(* IEC 61131-3 sources: nautilus/examples/remote-fleet/scada, 2 files *)

(* ---- sparkplug_types.st ---- *)
(*
  Generated by `naut sparkplug import` from the group's NBIRTH template
  definitions. Do not edit — re-run the import when a site's UDTs change.
  Group: Water
*)

TYPE
  Pump : STRUCT
    Run : BOOL;
    Fault : BOOL;
    SpeedHz : LREAL;
    SpeedSP : LREAL;
  END_STRUCT;
END_TYPE

(* Add the tags your program uses to its VAR_EXTERNAL block. The __Online,
   __Outages, __LastBirthMs and __Rebirth tags are synthesized by the driver:
   interlock on __Online before trusting a site's values, and pulse
   __Rebirth to force a resync. __Outages counts the times __Online went
   false.

VAR_EXTERNAL
  Booster1_DischargePress : LREAL;
  Booster1_FM1_FM1_FlowLps : LREAL;
  Booster1_FM1__Online : BOOL;
  Booster1_FM1__Outages : DINT;
  Booster1_Pump1 : Pump;
  Booster1_Pump1_SpeedSP : LREAL;
  Booster1_Pump2 : Pump;
  Booster1_Pump2_SpeedSP : LREAL;
  Booster1_SuctionPress : LREAL;
  Booster1_TankLevel : LREAL;
  Booster1__LastBirthMs : LINT;
  Booster1__Online : BOOL;
  Booster1__Outages : DINT;
  Booster1__Rebirth : BOOL;
  Well1_Pump1 : Pump;
  Well1_Pump1_SpeedSP : LREAL;
  Well1_WellLevel : LREAL;
  Well1__LastBirthMs : LINT;
  Well1__Online : BOOL;
  Well1__Outages : DINT;
  Well1__Rebirth : BOOL;
  Well2_Pump1 : Pump;
  Well2_Pump1_SpeedSP : LREAL;
  Well2_WellLevel : LREAL;
  Well2__LastBirthMs : LINT;
  Well2__Online : BOOL;
  Well2__Outages : DINT;
  Well2__Rebirth : BOOL;
END_VAR
*)

(* ---- fleet.st ---- *)
(* fleet.st — rollups over the whole consumed fleet, plus the plant's own
   local chlorine analyser. A site's data tag reads the zero of its type
   (quality notConnected) until the site first births, so __Online guards
   every one of them below: a never-birthed site must not count as a
   zero reading (nautilus.joyautomation.com/guides/sparkplug-host/). *)
PROGRAM Main
VAR_EXTERNAL
    Well1__Online     : BOOL;
    Well2__Online     : BOOL;
    Booster1__Online  : BOOL;
    Booster1_FM1__Online : BOOL;
    SitesOnline       : INT;

    Well1_Pump1       : Pump;
    Well2_Pump1       : Pump;
    Booster1_Pump1    : Pump;
    Booster1_Pump2    : Pump;
    AnyPumpRunning    : BOOL;

    Booster1_FM1_FM1_FlowLps : LREAL;
    SystemDemandLps   : LREAL;

    Booster1_TankLevel : LREAL;
    TankLevelPct       : LREAL;
    TankLowSP          : LREAL;
    TankLowAlm         : BOOL;

    CL1_ResidualPpm    : LREAL;
    ResidualLowSP      : LREAL;
    ChlorineResidualLowAlm : BOOL;
END_VAR

SitesOnline := 0;
IF Well1__Online THEN
    SitesOnline := SitesOnline + 1;
END_IF;
IF Well2__Online THEN
    SitesOnline := SitesOnline + 1;
END_IF;
IF Booster1__Online THEN
    SitesOnline := SitesOnline + 1;
END_IF;

AnyPumpRunning := (Well1__Online AND Well1_Pump1.Run)
    OR (Well2__Online AND Well2_Pump1.Run)
    OR (Booster1__Online AND (Booster1_Pump1.Run OR Booster1_Pump2.Run));

(* The system's own flow demand: Booster 1's discharge flow meter,
   guarded on ITS device's own online companion — a Modbus device
   attached to a Sparkplug node has its own __Online distinct from the
   node's. *)
IF Booster1_FM1__Online THEN
    SystemDemandLps := Booster1_FM1_FM1_FlowLps;
ELSE
    SystemDemandLps := 0.0;
END_IF;

(* The tank rollup — one site's reading, guarded the same way every other
   fleet value is. A dark Booster 1 reads as an empty tank, not a frozen
   last-known level: conservative, and consistent with "never trust a
   dead site's last value" everywhere else in this project. *)
IF Booster1__Online THEN
    TankLevelPct := Booster1_TankLevel;
ELSE
    TankLevelPct := 0.0;
END_IF;
TankLowAlm := TankLevelPct < TankLowSP;

(* The plant's own local device — no Sparkplug __Online to guard on; a
   disconnected Modbus source just holds its last-read value, same
   contract as every other field driver in this codebase. *)
ChlorineResidualLowAlm := CL1_ResidualPpm < ResidualLowSP;
END_PROGRAM
